Fanuc KAREL source: kd00040.KL

PROGRAM KD00040
%STACKSIZE=65535
%PRIORITY=65535
%NOLOCKGROUP
VAR
I : INTEGER
J : INTEGER
B : BOOLEAN
R : REAL
S : STRING[80]
-- UNRESOLVED DECLARATIONS (source type spelling not recovered)
-- PTH : TYPE_0x001F (type_u16=0x001F)
BEGIN
-- UNRESOLVED_PC line 11 opcodes [AD 32 22 9B 9B 9C 9C 37 2C] marker_code=0
END KD00040
